INTERFACE iRelay

PROPERTY PUBLIC IsSet : BOOL
GET
END_GET
END_PROPERTY

METHOD Reset
VAR_INPUT
END_VAR
END_METHOD

METHOD Set
VAR_INPUT
END_VAR
END_METHOD

END_INTERFACE

(* stored: Version 1.1.0.1
   Itf iRelay: Id {e3cfaf5b-d97f-49b8-86e4-4a18e56172f6}
   Property IsSet: Id {8a4b2fff-124d-4401-8d2b-2ab114f764de}
   Get Get: Id {23762f9c-c9d0-4857-8def-d07098c24431}
   Method Reset: Id {8832a2fe-12bf-40a0-9ba3-a21fe717fbe8}
   Method Set: Id {f9dfc50d-19c3-4d2f-9afa-e89c4ffba0a7} *)
